(* IEC 61131-3 sources: BODAS-HelloWorld/st/bodas_rc18_12_40/plc_logic/application/03_privatelibrary/datatypes/debugmanager, 3 files *)

(* ---- struc_dbgmgr-struc_DbgMgr.st ---- *)
(* --- Interface --- *)
TYPE struc_DbgMgr : STRUCT
		prm_struc  : struc_DbgMgrPrm;
		prv_struc  : struc_DbgMgrPrv;
		outp_struc : struc_DbgMgrOutp;
	END_STRUCT
END_TYPE

(* ---- struc_dbgmgroutp-struc_DbgMgrOutp.st ---- *)
(* --- Interface --- *)
TYPE struc_DbgMgrOutp : STRUCT
		flgStoreDataToNvmReq_l : BOOL; (* Flag TO store data TO NVM *)
	END_STRUCT
END_TYPE

(* ---- struc_dbgmgrprv-struc_DbgMgrPrv.st ---- *)
(* --- Interface --- *)
TYPE struc_DbgMgrPrv : STRUCT
		stErrDetn_u32           : UDINT; (* Status error detection *)
		flgStoreDataToNvmPrev_l : BOOL;  (* Flag TO store data TO NVM *)
	END_STRUCT
END_TYPE
